# EPICS autosave request: iocs/syringepump-ioc/db/ISCOController_settings.req
$(P)PressUnits
$(P)FlowUnits
$(P)OverpressAlarm
$(P)OverpressDisplay
$(P)UnderpressAlarm
$(P)UnderpressDisplay
$(P)UnderpressShutdown
$(P)OverflowAlarm
$(P)OverflowDisplay
$(P)OverflowShutdown
$(P)UnderflowAlarm
$(P)UnderflowDisplay
$(P)UnderflowShutdown
$(P)AB:DeliverToPercent
$(P)CD:DeliverToPercent
$(P)AB:RefillToPercent
$(P)CD:RefillToPercent
$(P)AB:Independent
$(P)CD:Independent
$(P)AB:DeliverMode
$(P)CD:DeliverMode
$(P)AB:PressureMode
$(P)CD:PressureMode
$(P)AB:PressureMatch
$(P)CD:PressureMatch
